(* CODESYS project tcl_unittestlibrary.library
   Company: Red Rock Controls Limited
   Description: TestRunner added
   Version: 1.2.0.0
   Placeholder: tcl_UnitTestLibrary
   Author: Roger Christopher
   Title: tcl_UnitTestLibrary

Project tree, tasks and I/O mapping:
  libraries: Tc2_Standard, * (Beckhoff Automation GmbH); Tc2_System, * (Beckhoff Automation GmbH); Tc2_Utilities, * (Beckhoff Automation GmbH); Tc3_EventLogger, * (Beckhoff Automation GmbH); Tc3_Module, * (Beckhoff Automation GmbH); tcl_BaseClasses, * (Red Rock Controls Limited)
  Functions/
    function F_LogError [ST]
    function F_LogMessage [ST]
  Message Buffer/
    function block T_MessageBuffer [ST]: AddMessage, GetMessage, LogCritical, LogDebug, LogError, LogInfo, LogWarning
  POUs/
    program PB_UnitTests [ST]
    function block T_Test1 [ST]: RunTest
    function block T_Test2 [ST]: RunTest
    function block T_Test3 [ST]: RunTest
  String Utils/
    function FormatString1 [ST]
    function FormatString2 [ST]
    function FormatString3 [ST]
    function FormatStringEx1 [ST]
    function FormatStringEx2 [ST]
    function block StringSplitter [ST]: GetNext, GetRemainder, HasMore, Init
  Test Runner/
    data type E_TestStatus
    data type ST_TestStatus
    function block T_TestRunner [ST]: AddTest, ClearTests, CyclicUpdate
  Unit Test/
    interface I_UnitTest: Init, RunTest, Completed, ElapsedTime, Enabled, Name, TestStatus
    function block T_UnitTestBase [ST]: AssertEquals_ANY, AssertEquals_BLOB, AssertEquals_BOOL, AssertEquals_BYTE, AssertEquals_DINT, AssertEquals_INT, AssertEquals_Interface, AssertEquals_LINT, AssertEquals_LREAL, AssertEquals_PVOID, AssertEquals_REAL, AssertEquals_STRING, AssertEquals_UDINT, AssertEquals_UINT, AssertEquals_ULINT, AssertEquals_USINT, AssertIsFalse, AssertIsTrue, Fail, FB_init, Init, RunTest, Completed, ElapsedTime, Enabled, Name, TestStatus
  Version/
    global variables Global_Version
  global variables Globals
*)

// Test Runner/E_TestStatus
{attribute 'qualified_only'}
{attribute 'strict'}
TYPE E_TestStatus :
(
	Unknown := 0,
	Running,
	Passed,
	Failed
);
END_TYPE

// Test Runner/ST_TestStatus
TYPE
    ST_TestStatus :
    STRUCT
        Name    : T_MaxString;
        Status  : E_TestStatus;
        Enabled : BOOL := TRUE;
    END_STRUCT
END_TYPE

// Version/Global_Version
{attribute 'TcGenerated'}
{attribute 'no-analysis'}
{attribute 'linkalways'}
// This function has been automatically generated from the project information.
VAR_GLOBAL CONSTANT
	{attribute 'const_non_replaced'}
	stLibVersion_tcl_UnitTestLibrary : ST_LibVersion := (iMajor := 1, iMinor := 2, iBuild := 0, iRevision := 0, nFlags := 0, sVersion := '1.2.0.0');
END_VAR

// Globals
//{attribute 'qualified_only'}
VAR_GLOBAL
//	DefaultLogger : T_MessageBuffer;
END_VAR

// Functions/F_LogError
FUNCTION INTERNAL F_LogError : BOOL
VAR_INPUT
    Source  : T_MaxString;
    Message : T_MaxString;
END_VAR
VAR
END_VAR

ADSLOGSTR(msgCtrlMask := ADSLOG_MSGTYPE_STRING OR ADSLOG_MSGTYPE_ERROR OR ADSLOG_MSGTYPE_LOG,
          msgFmtStr   := FormatStringEx2('%s : %s', Source, Message),
          strArg      := '');

END_FUNCTION

// String Utils/FormatStringEx2
{attribute 'hide'}
FUNCTION INTERNAL FormatStringEx2 : T_MaxString
VAR_INPUT
	Format	: T_MaxString;
	arg1	: T_MaxString;
	arg2	: T_MaxString;
END_VAR
VAR
    FB_FormatString1 : FB_FormatString;
END_VAR

FB_FormatString1(sFormat := Format,
                 arg1    := F_STRING(arg1),
                 arg2    := F_STRING(arg2),
                 arg3    :=,
                 arg4    :=,
                 arg5    :=,
                 arg6    :=,
                 arg7    :=,
                 arg8    :=,
                 arg9    :=,
                 arg10   :=,
                 bError  =>,
                 nErrId  =>,
                 sOut    => FormatStringEx2);

END_FUNCTION

// Functions/F_LogMessage
FUNCTION INTERNAL F_LogMessage : BOOL
VAR_INPUT
    Source  : T_MaxString;
    Message : T_MaxString;
END_VAR
VAR
END_VAR

ADSLOGSTR(msgCtrlMask := ADSLOG_MSGTYPE_STRING OR ADSLOG_MSGTYPE_HINT OR ADSLOG_MSGTYPE_LOG,
          msgFmtStr   := FormatStringEx2('%s : %s', Source, Message),
          strArg      := '');

END_FUNCTION

// Message Buffer/T_MessageBuffer
FUNCTION_BLOCK T_MessageBuffer
VAR
	MessageCount : UINT;
	Messages : ARRAY[0..MaxMessages] OF T_MaxString;
END_VAR
VAR CONSTANT
	MaxMessages : UINT := 99;
END_VAR

METHOD AddMessage : BOOL
VAR_INPUT
	Message : T_MaxString;
END_VAR
IF MessageCount < MaxMessages THEN
	Messages[MessageCount] := Message;
	F_Inc(MessageCount);
	AddMessage := TRUE;
END_IF
END_METHOD

METHOD GetMessage : T_MaxString
VAR_INPUT
END_VAR
IF MessageCount > 0 THEN
    GetMessage := Messages[0];
	F_Dec(MessageCount);		
	IF MessageCount > 0 THEN
		MEMMOVE(destAddr :=ADR(Messages[0]),
				srcAddr  :=ADR(Messages[1]),
				n        :=MessageCount * SIZEOF(T_MaxString));
	END_IF
END_IF
END_METHOD

METHOD LogCritical
VAR_INPUT
	Source	: T_MaxString;
	Message	: T_MaxString;
END_VAR
AddMessage(Message);
END_METHOD

METHOD LogDebug
VAR_INPUT
	Source	: T_MaxString;
	Message	: T_MaxString;
END_VAR
AddMessage(Message);
END_METHOD

METHOD LogError
VAR_INPUT
	Source	: T_MaxString;
	Message	: T_MaxString;
END_VAR
AddMessage(Message);
END_METHOD

METHOD LogInfo
VAR_INPUT
	Source	: T_MaxString;
	Message	: T_MaxString;
END_VAR
AddMessage(Message);
END_METHOD

METHOD LogWarning
VAR_INPUT
	Source	: T_MaxString;
	Message	: T_MaxString;
END_VAR
AddMessage(Message);
END_METHOD

END_FUNCTION_BLOCK

// POUs/PB_UnitTests
PROGRAM PB_UnitTests
VAR
	TestRunner : T_TestRunner;
	
	Test1 : T_Test1;
	Test2 : T_Test2;
	Test3 : T_Test3;
	
	Init : BOOL := TRUE;
	
END_VAR

IF Init THEN
	Init := FALSE;
	TestRunner.AddTest(Test1);
	TestRunner.AddTest(Test2);
	TestRunner.AddTest(Test3);
END_IF

TestRunner.CyclicUpdate();

END_PROGRAM

// Test Runner/T_TestRunner
FUNCTION_BLOCK T_TestRunner // TODO - remove TestStatus, move contents into T_UnitTestBase
VAR
    TaskTime          : LREAL;
    RunTests          : BOOL;
    Abort             : BOOL;
    EnableAllTests    : BOOL;
    DisableAllTests   : BOOL;
    Tests             : ARRAY[0..MaxTests] OF I_UnitTest;
    TestCount         : INT;
    FailedCount       : INT;
    CompletedCount    : INT;
    DisabledCount     : INT;
    CurrentTestNumber : INT;
    i                 : INT;
    TestsCompleted    : BOOL;
    SourceInfo        : FB_TcSourceInfo := (sName := 'Test Runner');

    State :
        (
        sInit,
        sInitialiseTests,
        sRunTests,
        sTestsCompleted);
    MessageBuffer : T_MessageBuffer;

END_VAR
VAR CONSTANT
    MaxTests : INT := 100;
END_VAR

METHOD AddTest : BOOL
VAR_INPUT
	Test : I_UnitTest;
END_VAR
IF State = sInit AND TestCount <= MaxTests THEN
    Tests[TestCount] := Test;
    F_Inc(TestCount);
    AddTest := TRUE;
END_IF
END_METHOD

METHOD ClearTests
VAR_INPUT
END_VAR
IF State = sInit THEN
    FOR i := 0 TO MaxTests DO
        Tests[i] := 0;
    END_FOR
    TestCount      := 0;
    FailedCount    := 0;
    CompletedCount := 0;
    DisabledCount  := 0;
	TestsCompleted := FALSE;
END_IF
END_METHOD

METHOD CyclicUpdate
VAR_INST
    RisingEdge1 : T_RisingEdge;
END_VAR
IF TaskTime = 0 THEN
    TaskTime := F_TaskTime();
END_IF

CASE State OF
    sInit:
        IF F_ReadFlag(RunTests) THEN
            IF TestCount > 0 AND TestCount <= MaxTests THEN
                State := sInitialiseTests;
            END_IF
        END_IF

        IF F_ReadFlag(EnableAllTests) AND TestCount > 0 THEN
            FOR i := 0 TO TestCount - 1 DO
                Tests[i].Enabled := TRUE;
            END_FOR
        END_IF

        IF F_ReadFlag(DisableAllTests) AND TestCount > 0 THEN
            FOR i := 0 TO TestCount - 1 DO
                Tests[i].Enabled := FALSE;
            END_FOR
        END_IF

    sInitialiseTests:
        TestsCompleted := FALSE;
        FailedCount    := 0;
        CompletedCount := 0;
        DisabledCount  := 0;
        FOR i := 0 TO TestCount - 1 DO
            IF Tests[i] <> 0 THEN
                Tests[i].Init();
            END_IF
        END_FOR
        CurrentTestNumber := 0;
        State             := sRunTests;

    sRunTests:
        IF F_ReadFlag(Abort) THEN
            tcl_BaseClasses.DefaultLogger.LogWarning(SourceInfo, 'Testing aborted');
            State := sTestsCompleted;
        ELSIF CurrentTestNumber >= TestCount THEN
            State := sTestsCompleted;
        ELSE
            IF Tests[CurrentTestNumber] = 0 THEN
                F_Inc(CurrentTestNumber);

            ELSIF NOT Tests[CurrentTestNumber].Enabled THEN
                F_Inc(DisabledCount);
                F_Inc(CurrentTestNumber);

            ELSIF Tests[CurrentTestNumber].Completed THEN
                IF Tests[CurrentTestNumber].TestStatus = E_TestStatus.Failed THEN
                    F_Inc(FailedCount);
                ELSE
                    Tests[CurrentTestNumber].TestStatus := E_TestStatus.Passed;
                END_IF
                F_Inc(CurrentTestNumber);
                F_Inc(CompletedCount);

            ELSE
                Tests[CurrentTestNumber].TestStatus  := E_TestStatus.Running;
                Tests[CurrentTestNumber].ElapsedTime := Tests[CurrentTestNumber].ElapsedTime + TaskTime;
                Tests[CurrentTestNumber].RunTest();

            END_IF
        END_IF

    sTestsCompleted:
        TestsCompleted := TRUE;
        tcl_BaseClasses.DefaultLogger.LogInfo(SourceInfo, FormatString2('%d tests completed, %d tests failed', F_INT(CompletedCount), F_INT(FailedCount)));
        CurrentTestNumber := -1;
        State             := sInit;

END_CASE
END_METHOD

END_FUNCTION_BLOCK

// Unit Test/T_UnitTestBase
{attribute 'reflection'}
FUNCTION_BLOCK ABSTRACT T_UnitTestBase
VAR
    {attribute 'instance-path'}
    {attribute 'no_init'}
    {attribute 'analysis' := '-33'} // Inhibit unused variable warning
    InstanceName : T_MaxString;     // Initialised with the instance name

    Project    : T_MaxString;
    Plc        : T_MaxString;
    TestName   : T_MaxString;
    SourceInfo : FB_TcSourceInfo := (sName := 'Unknown');

    _ElapsedTime : LREAL;
    _TestStatus  : E_TestStatus;
    _Enabled     : BOOL := TRUE;
	_Completed   : BOOL;
    State        : INT;

END_VAR

METHOD PROTECTED AssertEquals_ANY : BOOL
VAR_INPUT
    Expected : ANY;
    Actual   : ANY;
    Message  : T_MaxString;
END_VAR
VAR
    ComparisonResult : DINT;
END_VAR
ComparisonResult := MEMCMP(pBuf1 := Expected.pValue,
                           pBuf2 := Actual.pValue,
                           n     := DINT_TO_UDINT(Actual.diSize));

IF Expected.TypeClass <> Actual.TypeClass THEN
    DefaultLogger.LogError(SourceInfo, FormatStringEx1('Assertion Failed - %s', Message));
	_TestStatus := E_TestStatus.Failed;
    RETURN;

ELSIF Expected.diSize <> Actual.diSize THEN
    DefaultLogger.LogError(SourceInfo, FormatStringEx1('Assertion Failed - %s', Message));
	_TestStatus := E_TestStatus.Failed;
    RETURN;

ELSIF ComparisonResult <> 0 THEN
    DefaultLogger.LogError(SourceInfo, FormatStringEx1('Assertion Failed - %s', Message));
	_TestStatus := E_TestStatus.Failed;
    RETURN;
END_IF

AssertEquals_ANY := TRUE;
END_METHOD

METHOD AssertEquals_BLOB : BOOL
VAR_INPUT
    Expected : ANY;
    Actual   : ANY;
    Message  : T_MaxString;
END_VAR
IF
    Expected.diSize <> Actual.diSize
THEN
    tcl_BaseClasses.DefaultLogger.LogError(SourceInfo,
                           FormatString1('%s: Sizes differ',
                                         F_STRING(Message)));
	_TestStatus := E_TestStatus.Failed;
    RETURN;

ELSIF
    Expected.TypeClass <> Actual.TypeClass
THEN
    tcl_BaseClasses.DefaultLogger.LogError(SourceInfo,
                           FormatString1('%s: Type classes differ',
                                         F_STRING(Message)));
	_TestStatus := E_TestStatus.Failed;
    RETURN;

ELSIF
    MEMCMP(pBuf1 := Expected.pValue, // TODO - convert to function
           pBuf2 := Actual.pValue,
           n     := DINT_TO_UDINT(Actual.diSize)) <>  0
THEN
    tcl_BaseClasses.DefaultLogger.LogError(SourceInfo,
                           FormatString1('%s: Contents differ',
                                         F_STRING(Message)));
	_TestStatus := E_TestStatus.Failed;
    RETURN;
ELSE
    AssertEquals_BLOB := TRUE;
END_IF
END_METHOD

METHOD PROTECTED AssertEquals_BOOL : BOOL
VAR_INPUT
    Expected : BOOL;
    Actual   : BOOL;
    Message  : T_MaxString;
END_VAR
VAR
    ExpectedAsString : STRING;
    ActualAsString   : STRING;
END_VAR
IF Expected <> Actual THEN
    ExpectedAsString := BOOL_TO_STRING(Expected);
    ActualAsString   := BOOL_TO_STRING(Actual);
    tcl_BaseClasses.DefaultLogger.LogError(SourceInfo,
                           FormatString3('%s: expected=%s, actual=%s',
                                         F_STRING(Message),
                                         F_STRINGEX(ExpectedAsString),
                                         F_STRINGEX(ActualAsString)));
	_TestStatus := E_TestStatus.Failed;
    RETURN;
END_IF

AssertEquals_BOOL := TRUE;
END_METHOD

METHOD PROTECTED AssertEquals_BYTE : BOOL
VAR_INPUT
    Expected : BYTE;
    Actual   : BYTE;
    Message  : T_MaxString;
END_VAR
IF Expected <> Actual THEN
    tcl_BaseClasses.DefaultLogger.LogError(SourceInfo,
                           FormatString3('%s: expected=0x%.2X, actual=0x%.2X',
                                         F_STRING(Message),
                                         F_BYTE(Expected),
                                         F_BYTE(Actual)));
	_TestStatus := E_TestStatus.Failed;
    RETURN;
END_IF

AssertEquals_BYTE := TRUE;
END_METHOD

METHOD PROTECTED AssertEquals_DINT : BOOL
VAR_INPUT
    Expected : DINT;
    Actual   : DINT;
    Message  : T_MaxString;
END_VAR
IF Expected <> Actual THEN
    tcl_BaseClasses.DefaultLogger.LogError(SourceInfo,
                           FormatString3('%s: expected=%d, actual=%d',
                                         F_STRING(Message),
                                         F_DINT(Expected),
                                         F_DINT(Actual)));
	_TestStatus := E_TestStatus.Failed;
    RETURN;
END_IF

AssertEquals_DINT := TRUE;
END_METHOD

METHOD PROTECTED AssertEquals_INT : BOOL
VAR_INPUT
    Expected : INT;
    Actual   : INT;
    Message  : T_MaxString;
END_VAR
IF Expected <> Actual THEN
    tcl_BaseClasses.DefaultLogger.LogError(SourceInfo,
                           FormatString3('Failed - %s: expected=%d, actual=%d',
                                         F_STRING(Message),
                                         F_INT(Expected),
                                         F_INT(Actual)));
	_TestStatus := E_TestStatus.Failed;
    RETURN;
END_IF

AssertEquals_INT := TRUE;
END_METHOD

METHOD PROTECTED AssertEquals_Interface : BOOL
VAR_INPUT
    Expected : __SYSTEM.IQueryInterface;
    Actual   : __SYSTEM.IQueryInterface;
    Message  : T_MaxString;
END_VAR
IF Expected <> Actual THEN
    tcl_BaseClasses.DefaultLogger.LogError(SourceInfo,
                           FormatString1('%s',
                                         F_STRING(Message)));
	_TestStatus := E_TestStatus.Failed;
    RETURN;
END_IF

AssertEquals_Interface := TRUE;
END_METHOD

METHOD PROTECTED AssertEquals_LINT : BOOL
VAR_INPUT
    Expected : LINT;
    Actual   : LINT;
    Message  : T_MaxString;
END_VAR
IF Expected <> Actual THEN
    tcl_BaseClasses.DefaultLogger.LogError(SourceInfo,
                           FormatString3('%s: expected=%d, actual=%d',
                                         F_STRING(Message),
                                         F_LINT(Expected),
                                         F_LINT(Actual)));
	_TestStatus := E_TestStatus.Failed;
    RETURN;
END_IF

AssertEquals_LINT := TRUE;
END_METHOD

METHOD PROTECTED AssertEquals_LREAL : BOOL
VAR_INPUT
    Expected : LREAL;
    Actual   : LREAL;
    Delta    : LREAL;
    Message  : T_MaxString;
END_VAR
IF ABS(Expected - Actual) > Delta THEN
    tcl_BaseClasses.DefaultLogger.LogError(SourceInfo,
                           FormatString3('%s: expected= %.3f, actual= %.3f',
                                         F_STRING(Message),
                                         F_LREAL(Expected),
                                         F_LREAL(Actual)));
	_TestStatus := E_TestStatus.Failed;
    RETURN;
END_IF

AssertEquals_LREAL := TRUE;
END_METHOD

METHOD PROTECTED AssertEquals_PVOID : BOOL
VAR_INPUT
    Expected : PVOID;
    Actual   : PVOID;
    Message  : T_MaxString;
END_VAR
IF Expected <> Actual THEN
    tcl_BaseClasses.DefaultLogger.LogError(SourceInfo,
                           FormatString3('%s: expected=%d, actual=%d',
                                         F_STRING(Message),
                                         F_PVOID(Expected),
                                         F_PVOID(Actual)));
	_TestStatus := E_TestStatus.Failed;
    RETURN;
END_IF

AssertEquals_PVOID := TRUE;
END_METHOD

METHOD PROTECTED AssertEquals_REAL : BOOL
VAR_INPUT
    Expected : REAL;
    Actual   : REAL;
    Delta    : REAL;
    Message  : T_MaxString;
END_VAR
IF ABS(Expected - Actual) > Delta THEN
    tcl_BaseClasses.DefaultLogger.LogError(SourceInfo,
                           FormatString3('%s: expected=%.3f, actual=%.3f',
                                         F_STRING(Message),
                                         F_REAL(Expected),
                                         F_REAL(Actual)));
	_TestStatus := E_TestStatus.Failed;
    RETURN;
END_IF

AssertEquals_REAL := TRUE;
END_METHOD

METHOD PROTECTED AssertEquals_STRING : BOOL
VAR_INPUT
    Expected : T_MaxString;
    Actual   : T_MaxString;
    Message  : T_MaxString;
END_VAR
IF Expected <> Actual THEN
    tcl_BaseClasses.DefaultLogger.LogError(SourceInfo,
                           FormatString3('%s: expected=%s, actual=%s',
                                         F_STRING(Message),
                                         F_STRING(Expected),
                                         F_STRING(Actual)));
	_TestStatus := E_TestStatus.Failed;
    RETURN;
END_IF

AssertEquals_STRING := TRUE;
END_METHOD

METHOD PROTECTED AssertEquals_UDINT : BOOL
VAR_INPUT
    Expected : UDINT;
    Actual   : UDINT;
    Message  : T_MaxString;
END_VAR
IF Expected <> Actual THEN
    tcl_BaseClasses.DefaultLogger.LogError(SourceInfo,
                           FormatString3('%s: expected=%d, actual=%d',
                                         F_STRING(Message),
                                         F_UDINT(Expected),
                                         F_UDINT(Actual)));
	_TestStatus := E_TestStatus.Failed;
    RETURN;
END_IF

AssertEquals_UDINT := TRUE;
END_METHOD

METHOD PROTECTED AssertEquals_UINT : BOOL
VAR_INPUT
    Expected : UINT;
    Actual   : UINT;
    Message  : T_MaxString;
END_VAR
IF Expected <> Actual THEN
    tcl_BaseClasses.DefaultLogger.LogError(SourceInfo,
                           FormatString3('%s: expected=%d, actual=%d',
                                         F_STRING(Message),
                                         F_UINT(Expected),
                                         F_UINT(Actual)));
	_TestStatus := E_TestStatus.Failed;
    RETURN;
END_IF

AssertEquals_UINT := TRUE;
END_METHOD

METHOD PROTECTED AssertEquals_ULINT : BOOL
VAR_INPUT
    Expected : ULINT;
    Actual   : ULINT;
    Message  : T_MaxString;
END_VAR
IF Expected <> Actual THEN
    tcl_BaseClasses.DefaultLogger.LogError(SourceInfo,
                           FormatString3('%s: expected=%d, actual=%d',
                                         F_STRING(Message),
                                         F_ULINT(Expected),
                                         F_ULINT(Actual)));
	_TestStatus := E_TestStatus.Failed;
    RETURN;
END_IF

AssertEquals_ULINT := TRUE;
END_METHOD

METHOD PROTECTED AssertEquals_USINT : BOOL
VAR_INPUT
    Expected : USINT;
    Actual   : USINT;
    Message  : T_MaxString;
END_VAR
IF Expected <> Actual THEN
    tcl_BaseClasses.DefaultLogger.LogError(SourceInfo,
                           FormatString3('%s: expected=%d, actual=%d',
                                         F_STRING(Message),
                                         F_USINT(Expected),
                                         F_USINT(Actual)));
	_TestStatus := E_TestStatus.Failed;
    RETURN;
END_IF

AssertEquals_USINT := TRUE;
END_METHOD

METHOD PROTECTED AssertIsFalse : BOOL
VAR_INPUT
    Condition : BOOL;
    Message   : T_MaxString;
END_VAR
IF Condition THEN
    tcl_BaseClasses.DefaultLogger.LogError(SourceInfo,
                           FormatString1('%s: expected=FALSE, actual=TRUE',
                                         F_STRING(Message)));
	_TestStatus := E_TestStatus.Failed;
    RETURN;
END_IF

AssertIsFalse := TRUE;
END_METHOD

METHOD PROTECTED AssertIsTrue : BOOL
VAR_INPUT
    Condition : BOOL;
    Message   : T_MaxString;
END_VAR
IF NOT Condition THEN
    tcl_BaseClasses.DefaultLogger.LogError(SourceInfo,
                           FormatString1('%s: expected=TRUE, actual=FALSE',
                                         F_STRING(Message)));
	_TestStatus := E_TestStatus.Failed;
    RETURN;
END_IF

AssertIsTrue := TRUE;
END_METHOD

METHOD Fail
VAR_INPUT
    Message : T_MaxString;
END_VAR
tcl_BaseClasses.DefaultLogger.LogError(SourceInfo, FormatString1('Test Failure - %s', F_STRING(Message)));
_TestStatus := E_TestStatus.Failed;
END_METHOD

METHOD FB_init : BOOL
VAR_INPUT
	bInitRetains : BOOL; // if TRUE, the retain variables are initialized (warm start / cold start)
	bInCopyCode : BOOL;  // if TRUE, the instance afterwards gets moved into the copy code (online change)
END_VAR
VAR
	StringSplitter : StringSplitter;
END_VAR
StringSplitter.Init(Str    := InstanceName,
                    Delim1 := '.',
                    Delim2 := '');

IF StringSplitter.HasMore() THEN
    Project := StringSplitter.GetNext();
    Plc     := StringSplitter.GetNext();
END_IF

WHILE StringSplitter.HasMore() DO
    TestName := StringSplitter.GetNext(); // gets last chunk, which is Test Name
END_WHILE

SourceInfo.sName := TestName;

Init();
END_METHOD

METHOD Init
VAR_INPUT
END_VAR
_ElapsedTime := 0.0;
_TestStatus := E_TestStatus.Unknown;
_Completed := FALSE;State        := 0;
END_METHOD

{attribute 'analysis' := '-33'} // inhibit unused variable warning
METHOD ABSTRACT RunTest
END_METHOD

PROPERTY Completed : BOOL
GET
Completed := _Completed;
END_GET
END_PROPERTY

PROPERTY ElapsedTime : LREAL
GET
ElapsedTime := _ElapsedTime;
END_GET
SET
_ElapsedTime := ElapsedTime;
END_SET
END_PROPERTY

PROPERTY Enabled : BOOL
GET
Enabled := _Enabled;
END_GET
SET
_Enabled := Enabled;
END_SET
END_PROPERTY

{attribute 'monitoring' := 'call'}
PROPERTY Name : T_MaxString
GET
Name := TestName;
END_GET
END_PROPERTY

PROPERTY TestStatus : E_TestStatus
GET
TestStatus := _TestStatus;
END_GET
SET
_TestStatus := TestStatus;
END_SET
END_PROPERTY

END_FUNCTION_BLOCK

// String Utils/FormatStringEx1
{attribute 'hide'}
FUNCTION INTERNAL FormatStringEx1 : T_MaxString
VAR_INPUT
	Format	: T_MaxString;
	arg1	: T_MaxString;
END_VAR
VAR
    FB_FormatString1 : FB_FormatString;
END_VAR


FB_FormatString1(sFormat := Format,
                 arg1    := F_STRING(arg1),
                 arg2    :=,
                 arg3    :=,
                 arg4    :=,
                 arg5    :=,
                 arg6    :=,
                 arg7    :=,
                 arg8    :=,
                 arg9    :=,
                 arg10   :=,
                 bError  =>,
                 nErrId  =>,
                 sOut    => FormatStringEx1);

END_FUNCTION

// String Utils/FormatString1
{attribute 'hide'}
FUNCTION INTERNAL FormatString1 : T_MaxString
VAR_INPUT
	Format	: T_MaxString;
	arg1	: T_Arg;
END_VAR
VAR
    FB_FormatString1 : FB_FormatString;
END_VAR

FB_FormatString1(sFormat := Format,
                 arg1    := arg1,
                 arg2    :=,
                 arg3    :=,
                 arg4    :=,
                 arg5    :=,
                 arg6    :=,
                 arg7    :=,
                 arg8    :=,
                 arg9    :=,
                 arg10   :=,
                 bError  =>,
                 nErrId  =>,
                 sOut    => FormatString1);

END_FUNCTION

// String Utils/FormatString3
{attribute 'hide'}
FUNCTION INTERNAL FormatString3 : T_MaxString
VAR_INPUT
	Format	: T_MaxString;
	arg1	: T_Arg;
	arg2	: T_Arg;
	arg3	: T_Arg;
END_VAR
VAR
    FB_FormatString1 : FB_FormatString;
END_VAR

FB_FormatString1(sFormat := Format,
                 arg1    := arg1,
                 arg2    := arg2,
                 arg3    := arg3,
                 arg4    :=,
                 arg5    :=,
                 arg6    :=,
                 arg7    :=,
                 arg8    :=,
                 arg9    :=,
                 arg10   :=,
                 bError  =>,
                 nErrId  =>,
                 sOut    => FormatString3);

END_FUNCTION

// String Utils/StringSplitter
{attribute 'hide'}
FUNCTION_BLOCK INTERNAL StringSplitter
VAR
	SubjectString : TC2_SYSTEM.T_MaxString;
	Delimiter : STRING;
	Delimiter1 : STRING;
	Delimiter2 : STRING;
	NextDelimiterPosition : INT;
	NextDelimiter1Position : INT;
	NextDelimiter2Position : INT;
END_VAR

METHOD GetNext : STRING(255)
VAR_INPUT
END_VAR
VAR
	RemainingLength: INT;
END_VAR
NextDelimiter1Position := FIND(SubjectString , Delimiter1);
NextDelimiter2Position := FIND(SubjectString , Delimiter2);

IF NextDelimiter1Position = 0 THEN
    // use Delimiter 2 position , even if zero...
    NextDelimiterPosition := NextDelimiter2Position;
    Delimiter := Delimiter2;
    
ELSIF NextDelimiter2Position = 0 THEN
    // use Delimiter 1 position , non-zero...
    NextDelimiterPosition := NextDelimiter1Position;
    Delimiter := Delimiter1;

ELSE
    // Both delimters found - use the one nearest the start of the string...
    IF NextDelimiter1Position < NextDelimiter2Position THEN
        NextDelimiterPosition := NextDelimiter1Position;
        Delimiter := Delimiter1;
    ELSE
        NextDelimiterPosition := NextDelimiter2Position;
        Delimiter := Delimiter2;
	END_IF
END_IF

IF NextDelimiterPosition > 0 THEN // delimitter found
    
    // extract next sub-string
	GetNext := LEFT(SubjectString,NextDelimiterPosition - 1);
    
    // remove sub-string from subject string
	RemainingLength := LEN(SubjectString) - NextDelimiterPosition - LEN(Delimiter) + 1;
	SubjectString := RIGHT(SubjectString,RemainingLength);
    
//    // strip any delimitters from front of remaining string
//    WHILE FIND(SubjectString,Delimiter1) = 1 DO
//        SubjectString := RIGHT(SubjectString,LEN(SubjectString) - LEN(Delimiter1));
//	END_WHILE
//    WHILE FIND(SubjectString,Delimiter2) = 1 DO
//        SubjectString := RIGHT(SubjectString,LEN(SubjectString) - LEN(Delimiter2));
//	END_WHILE
ELSE
	GetNext := SubjectString; // return what is left
	SubjectString := '';
END_IF
END_METHOD

METHOD GetRemainder : STRING(255)
GetRemainder := SubjectString; // return what is left
SubjectString := '';
END_METHOD

METHOD HasMore : BOOL
VAR_INPUT
END_VAR
HasMore := SubjectString <> '';
END_METHOD

METHOD Init
VAR_INPUT
		Str : TC2_SYSTEM.T_MaxString;
		Delim1 : STRING;
		Delim2 : STRING;
END_VAR
SubjectString := Str;
NextDelimiterPosition := 0;
Delimiter1 := Delim1;
Delimiter2 := Delim2;
END_METHOD

END_FUNCTION_BLOCK

// Unit Test/I_UnitTest
INTERFACE I_UnitTest

METHOD Init
VAR

END_VAR
END_METHOD

METHOD ABSTRACT RunTest
END_METHOD

PROPERTY Completed : BOOL
GET
END_GET
END_PROPERTY

PROPERTY ElapsedTime : LREAL
GET
END_GET
SET
END_SET
END_PROPERTY

{attribute 'monitoring' := 'call'}
PROPERTY Enabled : BOOL
GET
END_GET
SET
END_SET
END_PROPERTY

{attribute 'monitoring' := 'call'}
PROPERTY Name : T_MaxString
GET
END_GET
END_PROPERTY

{attribute 'monitoring' := 'call'}
PROPERTY TestStatus : E_TestStatus
GET
END_GET
SET
END_SET
END_PROPERTY

END_INTERFACE

// String Utils/FormatString2
{attribute 'hide'}
FUNCTION INTERNAL FormatString2 : T_MaxString
VAR_INPUT
	Format	: T_MaxString;
	arg1	: T_Arg;
	arg2	: T_Arg;
END_VAR
VAR
    FB_FormatString1 : FB_FormatString;
END_VAR

FB_FormatString1(sFormat := Format,
                 arg1    := arg1,
                 arg2    := arg2,
                 arg3    :=,
                 arg4    :=,
                 arg5    :=,
                 arg6    :=,
                 arg7    :=,
                 arg8    :=,
                 arg9    :=,
                 arg10   :=,
                 bError  =>,
                 nErrId  =>,
                 sOut    => FormatString2);

END_FUNCTION

// POUs/T_Test1
FUNCTION_BLOCK T_Test1 EXTENDS T_UnitTestBase IMPLEMENTS I_UnitTest
VAR
	Value : INT := 7;
END_VAR

{attribute 'analysis' := '-33'} // inhibit unused variable warning
METHOD  RunTest
VAR_INST
	OnTimer : T_OnTimer(PresetTime := 1.5);
END_VAR
CASE State OF
    0:
        OnTimer.Reset();
        Value := 5;
        F_Inc(State);
    1:
        AssertEquals_INT(Expected := 7, Actual := Value, Message := 'Value');
        F_Inc(State);

    2:
        IF OnTimer.Run() THEN
            _Completed := TRUE;
        END_IF

END_CASE
END_METHOD

END_FUNCTION_BLOCK

// POUs/T_Test2
FUNCTION_BLOCK T_Test2 EXTENDS T_UnitTestBase IMPLEMENTS I_UnitTest
VAR
	Value : INT := 7;
END_VAR

{attribute 'analysis' := '-33'} // inhibit unused variable warning
METHOD  RunTest
VAR_INST
	OnTimer : T_OnTimer(PresetTime := 1.0);
END_VAR
CASE State OF
    0:
        OnTimer.Reset();
        Value := 5;
        F_Inc(State);
    1:
        AssertEquals_INT(Expected := 7, Actual := Value, Message := 'Value');
        F_Inc(State);

    2:
        IF OnTimer.Run() THEN
            _Completed := TRUE;
        END_IF

END_CASE
END_METHOD

END_FUNCTION_BLOCK

// POUs/T_Test3
FUNCTION_BLOCK T_Test3 EXTENDS T_UnitTestBase IMPLEMENTS I_UnitTest
VAR
	Value : INT := 7;
END_VAR

{attribute 'analysis' := '-33'} // inhibit unused variable warning
METHOD  RunTest
VAR_INST
	OnTimer : T_OnTimer(PresetTime := 2.0);
END_VAR
CASE State OF
    0:
        OnTimer.Reset();
        F_Inc(State);
		
    1:
		Fail('Fail reason here');
        F_Inc(State);

    2:
        IF OnTimer.Run() THEN
            _Completed := TRUE;
        END_IF

END_CASE
END_METHOD

END_FUNCTION_BLOCK
